FUNCTION_BLOCK FB_Pump EXTENDS FB_Device
VAR_INPUT
	bRunReq : BOOL;   // program wants the pump running
END_VAR
VAR_OUTPUT
	bRunCmd : BOOL;   // contactor output
END_VAR

bRunCmd := bRunReq AND NOT bFault;

END_FUNCTION_BLOCK

(* stored: Version 1.1.0.1, ProductVersion 3.1.4026.12
   POU FB_Pump: Id {3a2b3c4d-0000-4000-8000-000000000002}, SpecialFunc None *)
